// TIA Portal V21 export
Screen "R05_BtnNav"  1024x768, Number=44, Template=Tpl
  ScreenLayer 
    Button "P_NavBtn" at 10,10 size 100x30  TextOff="BTN", TextOn="BTN"
      on Press: ActivateScreen(Screen name := Alarms, Object number := 0)
